(* IEC 61131-3 sources: Codesys-MCP-Server/examples/heatpump/st, 12 files *)

(* ---- E_HpState.st ---- *)
{attribute 'qualified_only'}
TYPE E_HpState :
(
	OFF := 0,
	STANDBY := 1,
	PREPUMP := 2,
	HEATING := 3,
	DHW := 4,
	POSTPUMP := 5,
	FAULT := 6
);
END_TYPE

(* ---- GVL_IO.st ---- *)
{attribute 'qualified_only'}
VAR_GLOBAL
	// --- Eingaenge (Analog, degC) ---
	rTempOutside  : REAL;   // Aussentemperatur
	rTempFlow     : REAL;   // Vorlauftemperatur
	rTempReturn   : REAL;   // Ruecklauftemperatur
	rTempDHW      : REAL;   // Warmwasser-Speicher
	rTempSource   : REAL;   // Quelle (Sole/Verdampfer)
	// --- Eingaenge (Digital) ---
	xHighPressure : BOOL;   // Hochdruckwaechter (TRUE=Stoerung)
	xLowPressure  : BOOL;   // Niederdruckwaechter (TRUE=Stoerung)
	xFlowSwitch   : BOOL;   // Stroemungswaechter (TRUE=Durchfluss ok)
	xDemand       : BOOL;   // Externe Heizanforderung / Thermostat
	xReset        : BOOL;   // Stoerungs-Quittierung
	// --- Ausgaenge (Digital) ---
	xCompressor   : BOOL;   // Verdichter-Schuetz
	xSourcePump   : BOOL;   // Quellenpumpe / Ventilator
	xSinkPump     : BOOL;   // Heizkreispumpe
	xValveDHW     : BOOL;   // 3-Wege-Ventil (TRUE=Warmwasser)
	xBackupHeater : BOOL;   // Elektro-Zusatzheizung
	xFaultLamp    : BOOL;   // Stoermeldeleuchte
END_VAR

(* ---- GVL_Param.st ---- *)
{attribute 'qualified_only'}
VAR_GLOBAL CONSTANT
	// Heizkurve: Vorlauf-Sollwert linear ueber Aussentemperatur
	rHC_OutMin  : REAL := -15.0;
	rHC_FlowMax : REAL := 45.0;
	rHC_OutMax  : REAL := 18.0;
	rHC_FlowMin : REAL := 25.0;
	rFlowHyst   : REAL := 3.0;
	// Warmwasser
	rDHW_Set    : REAL := 50.0;
	rDHW_Hyst   : REAL := 5.0;
	rDHW_Max    : REAL := 60.0;
	// Zusatzheizung (Bivalenzpunkt)
	rBackupOn   : REAL := -7.0;
	// Quelle
	rSourceMin  : REAL := -5.0;
	// Zeiten
	tPrePump    : TIME := T#30S;
	tPostPump   : TIME := T#60S;
	tMinRun     : TIME := T#5M;
	tMinOff     : TIME := T#5M;
	tFlowFault  : TIME := T#10S;
END_VAR

(* ---- FB_CompressorProtect.decl.st ---- *)
FUNCTION_BLOCK FB_CompressorProtect
VAR_INPUT
	xRequest : BOOL;
	tMinRun  : TIME;
	tMinOff  : TIME;
END_VAR
VAR_OUTPUT
	xCompressor : BOOL;
	xReady      : BOOL;
END_VAR
VAR
	tonRun : TON;
	tonOff : TON;
END_VAR

(* ---- FB_HeatCurve.decl.st ---- *)
FUNCTION_BLOCK FB_HeatCurve
VAR_INPUT
	rOutside : REAL;
	rOutMin  : REAL;
	rFlowMax : REAL;
	rOutMax  : REAL;
	rFlowMin : REAL;
END_VAR
VAR_OUTPUT
	rFlowSet : REAL;
END_VAR
VAR
	rX     : REAL;
	rSlope : REAL;
END_VAR

(* ---- FB_HeatPump.decl.st ---- *)
FUNCTION_BLOCK FB_HeatPump
VAR_INPUT
	rTempOutside  : REAL;
	rTempFlow     : REAL;
	rTempReturn   : REAL;
	rTempDHW      : REAL;
	rTempSource   : REAL;
	xHighPressure : BOOL;
	xLowPressure  : BOOL;
	xFlowSwitch   : BOOL;
	xDemand       : BOOL;
	xReset        : BOOL;
END_VAR
VAR_OUTPUT
	xCompressor   : BOOL;
	xSourcePump   : BOOL;
	xSinkPump     : BOOL;
	xValveDHW     : BOOL;
	xBackupHeater : BOOL;
	xFault        : BOOL;
	eState        : E_HpState;
	rFlowSet      : REAL;
END_VAR
VAR
	fbCurve   : FB_HeatCurve;
	fbHeatHy  : FB_Hysteresis;
	fbDhwHy   : FB_Hysteresis;
	fbProtect : FB_CompressorProtect;
	tonPre    : TON;
	tonPost   : TON;
	tonFlow   : TON;
	rtReset   : R_TRIG;
	xHeatReq  : BOOL;
	xDhwReq   : BOOL;
	xCompReq  : BOOL;
	xSafeOk   : BOOL;
END_VAR

(* ---- FB_Hysteresis.decl.st ---- *)
FUNCTION_BLOCK FB_Hysteresis
VAR_INPUT
	rActual : REAL;
	rSet    : REAL;
	rHyst   : REAL;
END_VAR
VAR_OUTPUT
	xDemand : BOOL;
END_VAR

(* ---- FB_CompressorProtect.impl.st ---- *)
// Taktschutz: Mindestlaufzeit + Mindeststillstand (Anti-Short-Cycle)
tonRun(IN := xCompressor, PT := tMinRun);
tonOff(IN := NOT xCompressor, PT := tMinOff);
xReady := tonOff.Q;
IF xCompressor THEN
	// laeuft: erst nach Mindestlaufzeit abschalten, wenn nicht mehr angefordert
	IF (NOT xRequest) AND tonRun.Q THEN
		xCompressor := FALSE;
	END_IF
ELSE
	// steht: erst nach Mindeststillstand und bei Anforderung starten
	IF xRequest AND xReady THEN
		xCompressor := TRUE;
	END_IF
END_IF

(* ---- FB_HeatCurve.impl.st ---- *)
// Aussentemperatur auf den Kurvenbereich begrenzen
rX := LIMIT(rOutMin, rOutside, rOutMax);
// lineare Interpolation zwischen (rOutMin,rFlowMax) und (rOutMax,rFlowMin)
IF (rOutMax - rOutMin) <> 0.0 THEN
	rSlope := (rFlowMin - rFlowMax) / (rOutMax - rOutMin);
	rFlowSet := rFlowMax + rSlope * (rX - rOutMin);
ELSE
	rFlowSet := rFlowMax;
END_IF

(* ---- FB_HeatPump.impl.st ---- *)
// === 1) Flanken und Zeiten (einmal pro Zyklus) ===
rtReset(CLK := xReset);
tonFlow(IN := xSinkPump AND NOT xFlowSwitch, PT := GVL_Param.tFlowFault);
tonPre(IN := (eState = E_HpState.PREPUMP), PT := GVL_Param.tPrePump);
tonPost(IN := (eState = E_HpState.POSTPUMP), PT := GVL_Param.tPostPump);

// === 2) Sicherheits-Sammelmeldung ===
xSafeOk := (NOT xHighPressure) AND (NOT xLowPressure)
           AND (NOT tonFlow.Q) AND (rTempSource > GVL_Param.rSourceMin);

// === 3) Sollwerte und Anforderungen ===
fbCurve(rOutside := rTempOutside,
        rOutMin := GVL_Param.rHC_OutMin, rFlowMax := GVL_Param.rHC_FlowMax,
        rOutMax := GVL_Param.rHC_OutMax, rFlowMin := GVL_Param.rHC_FlowMin);
rFlowSet := fbCurve.rFlowSet;

fbHeatHy(rActual := rTempFlow, rSet := rFlowSet, rHyst := GVL_Param.rFlowHyst);
xHeatReq := fbHeatHy.xDemand AND xDemand;

fbDhwHy(rActual := rTempDHW, rSet := GVL_Param.rDHW_Set, rHyst := GVL_Param.rDHW_Hyst);
xDhwReq := fbDhwHy.xDemand;

xCompReq := FALSE;

// === 4) Zustandsautomat ===
CASE eState OF

	E_HpState.OFF:
		xCompressor := FALSE; xSourcePump := FALSE; xSinkPump := FALSE;
		xBackupHeater := FALSE; xValveDHW := FALSE;
		IF xSafeOk THEN
			eState := E_HpState.STANDBY;
		END_IF

	E_HpState.STANDBY:
		xSourcePump := FALSE;
		xSinkPump := xHeatReq;
		xBackupHeater := FALSE;
		IF NOT xSafeOk THEN
			eState := E_HpState.FAULT;
		ELSIF xDhwReq OR xHeatReq THEN
			eState := E_HpState.PREPUMP;
		END_IF

	E_HpState.PREPUMP:
		xSourcePump := TRUE; xSinkPump := TRUE;
		xValveDHW := xDhwReq;
		IF NOT xSafeOk THEN
			eState := E_HpState.FAULT;
		ELSIF NOT (xDhwReq OR xHeatReq) THEN
			eState := E_HpState.POSTPUMP;
		ELSIF tonPre.Q THEN
			IF xDhwReq THEN
				eState := E_HpState.DHW;
			ELSE
				eState := E_HpState.HEATING;
			END_IF
		END_IF

	E_HpState.HEATING:
		xValveDHW := FALSE;
		xSourcePump := TRUE; xSinkPump := TRUE;
		xCompReq := xHeatReq;
		xBackupHeater := xHeatReq AND (rTempOutside <= GVL_Param.rBackupOn);
		IF NOT xSafeOk THEN
			eState := E_HpState.FAULT;
		ELSIF xDhwReq THEN
			eState := E_HpState.DHW;
		ELSIF NOT xHeatReq THEN
			eState := E_HpState.POSTPUMP;
		END_IF

	E_HpState.DHW:
		xValveDHW := TRUE;
		xSourcePump := TRUE; xSinkPump := TRUE;
		xCompReq := xDhwReq AND (rTempDHW < GVL_Param.rDHW_Max);
		xBackupHeater := FALSE;
		IF NOT xSafeOk THEN
			eState := E_HpState.FAULT;
		ELSIF NOT xDhwReq THEN
			IF xHeatReq THEN
				eState := E_HpState.HEATING;
			ELSE
				eState := E_HpState.POSTPUMP;
			END_IF
		END_IF

	E_HpState.POSTPUMP:
		xBackupHeater := FALSE;
		xSourcePump := TRUE; xSinkPump := TRUE;
		IF NOT xSafeOk THEN
			eState := E_HpState.FAULT;
		ELSIF xDhwReq OR xHeatReq THEN
			eState := E_HpState.PREPUMP;
		ELSIF tonPost.Q THEN
			eState := E_HpState.STANDBY;
		END_IF

	E_HpState.FAULT:
		xSourcePump := FALSE; xSinkPump := FALSE; xBackupHeater := FALSE;
		xFault := TRUE;
		IF rtReset.Q AND xSafeOk THEN
			xFault := FALSE;
			eState := E_HpState.OFF;
		END_IF

END_CASE

// === 5) Verdichter mit Taktschutz ===
xCompReq := xCompReq AND xSafeOk AND (eState <> E_HpState.FAULT);
fbProtect(xRequest := xCompReq, tMinRun := GVL_Param.tMinRun, tMinOff := GVL_Param.tMinOff);
xCompressor := fbProtect.xCompressor;

// === 6) Harte Sicherheits-Abschaltung hat immer Vorrang ===
IF NOT xSafeOk THEN
	xCompressor := FALSE;
	xBackupHeater := FALSE;
END_IF

(* ---- FB_Hysteresis.impl.st ---- *)
// Bistabile 2-Punkt-Hysterese: Anforderung EIN unter (Soll-Hyst), AUS bei Soll
IF rActual <= (rSet - rHyst) THEN
	xDemand := TRUE;
ELSIF rActual >= rSet THEN
	xDemand := FALSE;
END_IF

(* ---- PLC_PRG.decl.st ---- *)
PROGRAM PLC_PRG
VAR
	fbHeatPump : FB_HeatPump;
END_VAR
